(* Logix 5000 project; controller NWGG_Treater_Dayton vendor 1 type 14 code 238 rev 35.11; software revision 35.00; part 5 of 5 *)
(* tags used below, declared in another part *)
   Non_Water_Total_Chemical_Package : REAL;
   Total_Chemical_Package : REAL;
   Treater_Pump : Treater_Pump[50];
   Water : Analog_Gallon_Values;
(* Pumps, continued *)

ROUTINE Water   (* ladder *)
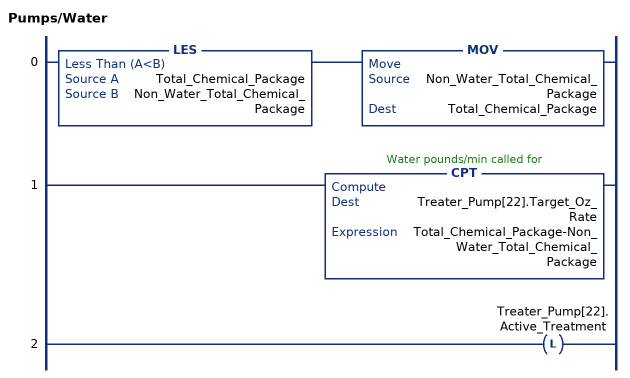
   0: LES(Total_Chemical_Package,Non_Water_Total_Chemical_Package)MOV(Non_Water_Total_Chemical_Package,Total_Chemical_Package);
   1: CPT(Treater_Pump[22].Target_Oz_Rate,Total_Chemical_Package-Non_Water_Total_Chemical_Package);
   2: OTL(Treater_Pump[22].Active_Treatment);
END_ROUTINE
END_PROGRAM

PROGRAM SafetyProgram   (* main routine MainRoutine, safety *)

ROUTINE MainRoutine   (* ladder *)
END_ROUTINE
END_PROGRAM
